Fanuc KAREL source: KT00938.KL

PROGRAM KT00938
%NOLOCKGROUP
VAR
  ENTRY: INTEGER
  PNAME: STRING[80]
  VNAME: STRING[80]
  STATUS: INTEGER
  VALUE: ARRAY[2] OF SHORT
BEGIN
  ENTRY = 0
  PNAME = ''
  VNAME = 'VALUE'
  VALUE[1] = 2
  GET_VAR(ENTRY, PNAME, VNAME, VALUE[1], STATUS)
END KT00938
